// TIA Portal V20 export
// export: Created 2026-11-12T11:17:33.9267401Z, ExportSetting WithDefaults, DisplayName Totally Integrated Automation Portal, DisplayVersion V20, DisplayName TIA Portal Openness, DisplayVersion V20, DisplayName TIA Portal Teamcenter Gateway, DisplayVersion V20, DisplayName TIA Portal Version Control Interface, DisplayVersion V20, DisplayName STEP 7 Professional, DisplayVersion V20, DisplayName STEP 7 CFC, DisplayVersion V20, DisplayName STEP 7 Safety, DisplayVersion V20, DisplayName WinCC Basic/Comfort/Advanced, DisplayVersion V20, DisplayName SIMATIC Visualization Architect, DisplayVersion V20, DisplayName WinCC Professional, DisplayVersion V20, DisplayName SIMATIC Visualization Architect, DisplayVersion V20, DisplayName WinCC Unified, DisplayVersion V20, DisplayName SIMATIC Visualization Architect, DisplayVersion V20
TYPE "UDT_Entradas_APP"
// stored: IsFailsafeCompliant false
   STRUCT
      Eje_z_arriba : Bool;
      Eje_z_abajo : Bool;
      Gripper_abierto : Bool;
      Almacen_izq_lleno : Bool;
      Almacen_dch_lleno : Bool;
      Eje_referenciado : Bool;
      Motion_complete : Bool;
      Ready : Bool;
   END_STRUCT;
END_TYPE
